// TIA Portal V21 export
// export: Created 2026-10-14T03:08:58.0952126Z, ExportSetting WithDefaults, DisplayName Totally Integrated Automation Portal, DisplayVersion V21, DisplayName STEP 7 Professional, DisplayVersion V21, DisplayName STEP 7 Safety, DisplayVersion V21, DisplayName Tech WebApplication, DisplayVersion V21, DisplayName WinCC Basic/Comfort/Advanced, DisplayVersion V21, DisplayName WinCC Unified, DisplayVersion V21
FUNCTION_BLOCK "FB_5_CIP_Simulation_Graph"   // FB7, GRAPH
VERSION : 0.1
// stored: AcknowledgeErrorsRequired true, AutoNumber true, GraphVersion 6.0, InitialValuesAcquisition false, IsIECCheckEnabled false, LanguageInNetworks LAD, LockOperatingMode false, PermanentILProcessingInMANMode false, SetENOAutomatically false, SkipSteps false, UDAEnableTagReadback false, WithAlarmHandling true
   // inherited from GRAPH_BASE
   VAR
      OFF_SQ_BASE : Bool;
   END_VAR
   VAR_INPUT
      OFF_SQ { ExternalAccessible := 'False'; ExternalVisible := 'False'; ExternalWritable := 'False'} : Bool := false;   // Turn sequence off
      INIT_SQ { ExternalAccessible := 'False'; ExternalVisible := 'False'; ExternalWritable := 'False'} : Bool := false;   // Set sequence to initial state
      ACK_EF { ExternalAccessible := 'False'; ExternalVisible := 'False'; ExternalWritable := 'False'} : Bool := false;   // Acknowledge all errors and faults
      S_PREV { ExternalAccessible := 'False'; ExternalVisible := 'False'; ExternalWritable := 'False'} : Bool := false;   // Output previous step in parameter S_NO
      S_NEXT { ExternalAccessible := 'False'; ExternalVisible := 'False'; ExternalWritable := 'False'} : Bool := false;   // Indicate next step in parameter S_NO
      SW_AUTO { ExternalAccessible := 'False'; ExternalVisible := 'False'; ExternalWritable := 'False'} : Bool := false;   // Automatic mode
      SW_TAP { ExternalAccessible := 'False'; ExternalVisible := 'False'; ExternalWritable := 'False'} : Bool := false;   // Semiautomatic/switch with transition
      SW_TOP { ExternalAccessible := 'False'; ExternalVisible := 'False'; ExternalWritable := 'False'} : Bool := false;   // Semiautomatic/ignore transition
      SW_MAN { ExternalAccessible := 'False'; ExternalVisible := 'False'; ExternalWritable := 'False'} : Bool := false;   // Manual mode
      S_SEL { ExternalAccessible := 'False'; ExternalVisible := 'False'; ExternalWritable := 'False'} : Int := 0;   // Select step to be output to S_NO
      S_ON { ExternalAccessible := 'False'; ExternalVisible := 'False'; ExternalWritable := 'False'} : Bool := false;   // Activate step indicated in S_NO
      S_OFF { ExternalAccessible := 'False'; ExternalVisible := 'False'; ExternalWritable := 'False'} : Bool := false;   // Disable step indicated in S_NO
      T_PUSH { ExternalAccessible := 'False'; ExternalVisible := 'False'; ExternalWritable := 'False'} : Bool := false;   // Enable transition to switch in semi automatic mode
   END_VAR
   VAR_OUTPUT
      S_NO { ExternalAccessible := 'False'; ExternalVisible := 'False'; ExternalWritable := 'False'} : Int := 0;   // Step number
      S_MORE { ExternalAccessible := 'False'; ExternalVisible := 'False'; ExternalWritable := 'False'} : Bool := false;   // More steps are available and can be shown in S_NO
      S_ACTIVE { ExternalAccessible := 'False'; ExternalVisible := 'False'; ExternalWritable := 'False'} : Bool := false;   // Step indicated in S_NO is active
      ERR_FLT { ExternalAccessible := 'False'; ExternalVisible := 'False'; ExternalWritable := 'False'} : Bool := false;   // Interlock or supervision group error
      AUTO_ON { ExternalAccessible := 'False'; ExternalVisible := 'False'; ExternalWritable := 'False'} : Bool := false;   // Automatic mode is active
      TAP_ON { ExternalAccessible := 'False'; ExternalVisible := 'False'; ExternalWritable := 'False'} : Bool := false;   // Semiautomatic mode/step with transition enabled
      TOP_ON { ExternalAccessible := 'False'; ExternalVisible := 'False'; ExternalWritable := 'False'} : Bool := false;   // Semiautomatic mode/ignore transition enabled
      MAN_ON { ExternalAccessible := 'False'; ExternalVisible := 'False'; ExternalWritable := 'False'} : Bool := false;   // Manual mode is active
   END_VAR
   VAR_IN_OUT
      cip : "typeCIP";
      stepInitial : Bool;   // Initial step is active
      step1Active : Bool;   // Step 1 is active
      step2Active : Bool;   // Step 2 is active
      step3Active : Bool;   // Step 3 is active
      step4Active : Bool;   // Step 4 is active
   END_VAR
   VAR
      statTemperature : Real;
      statConcentration : Real;
      statAbnomaly : Real;
   END_VAR
   VAR_TEMP
      tempRet : Int;
      tempRandomFlowrate : Int;
      tempRandomAbnomaly : Real;
   END_VAR
BEGIN
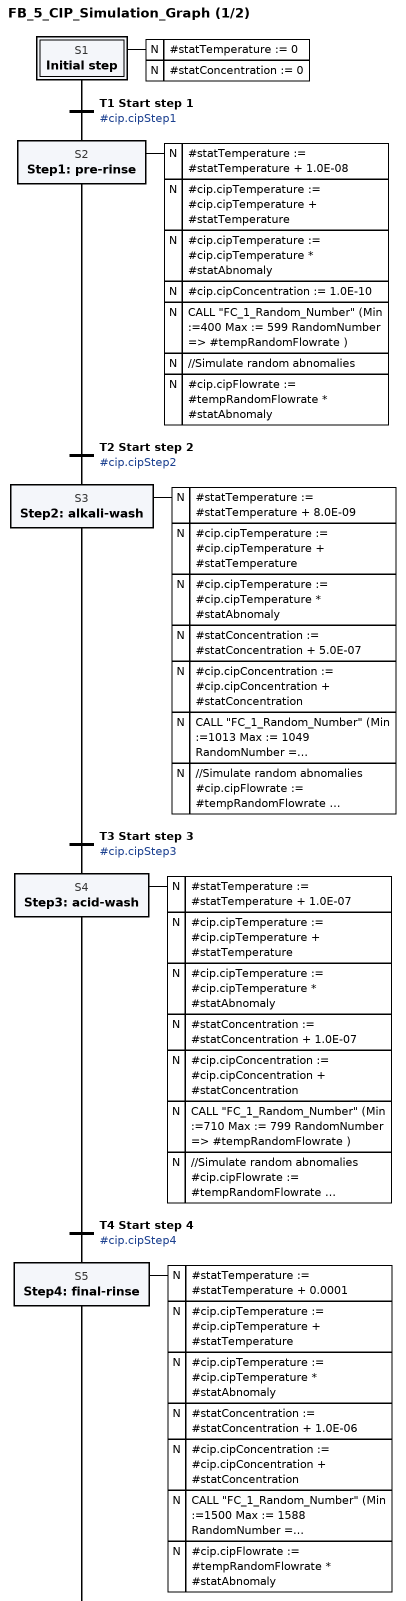
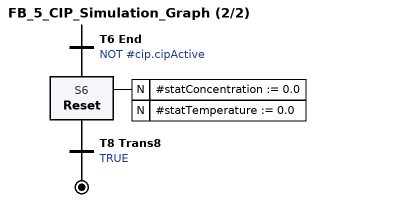
   // permanent pre-instructions
   NETWORK 1
   TITLE = Simulate random abnomalies
      "FC_1_Random_Number"(Min := 70, Max := 100, RandomNumber => #tempRandomAbnomaly);
      #statAbnomaly := #tempRandomAbnomaly / 100.0;

   // sequencer 1
   INITIAL_STEP "Initial step":   // S1, max time T#10S, warning time T#7S
              N    #statTemperature := 0
              N    #statConcentration := 0
   END_STEP
   TRANSITION "Start step 1" FROM "Initial step" TO "Step1: pre-rinse"   // T1
      := #cip.cipStep1;
   END_TRANSITION
   STEP "Step1: pre-rinse":   // S2, max time T#10S, warning time T#7S
              N    #statTemperature := #statTemperature + 1.0E-08
              N    #cip.cipTemperature := #cip.cipTemperature + #statTemperature
              N    #cip.cipTemperature := #cip.cipTemperature * #statAbnomaly
              N    #cip.cipConcentration := 1.0E-10
              N    CALL "FC_1_Random_Number"
                   (Min :=400
                   Max := 599
                   RandomNumber => #tempRandomFlowrate
                   )
                   //Simulate random abnomalies
              N    #cip.cipFlowrate := #tempRandomFlowrate * #statAbnomaly
   END_STEP
   TRANSITION "Start step 2" FROM "Step1: pre-rinse" TO "Step2: alkali-wash"   // T2
      := #cip.cipStep2;
   END_TRANSITION
   STEP "Step2: alkali-wash":   // S3, max time T#10S, warning time T#7S
              N    #statTemperature := #statTemperature + 8.0E-09
              N    #cip.cipTemperature := #cip.cipTemperature + #statTemperature
              N    #cip.cipTemperature := #cip.cipTemperature * #statAbnomaly
              N    #statConcentration := #statConcentration + 5.0E-07
              N    #cip.cipConcentration := #cip.cipConcentration + #statConcentration
              N    CALL "FC_1_Random_Number"
                   (Min :=1013
                   Max := 1049
                   RandomNumber => #tempRandomFlowrate
                   )
              N    //Simulate random abnomalies
                   #cip.cipFlowrate := #tempRandomFlowrate * #statAbnomaly
   END_STEP
   TRANSITION "Start step 3" FROM "Step2: alkali-wash" TO "Step3: acid-wash"   // T3
      := #cip.cipStep3;
   END_TRANSITION
   STEP "Step3: acid-wash":   // S4, max time T#10S, warning time T#7S
              N    #statTemperature := #statTemperature + 1.0E-07
              N    #cip.cipTemperature := #cip.cipTemperature + #statTemperature
              N    #cip.cipTemperature := #cip.cipTemperature * #statAbnomaly
              N    #statConcentration := #statConcentration + 1.0E-07
              N    #cip.cipConcentration := #cip.cipConcentration + #statConcentration
              N    CALL "FC_1_Random_Number"
                   (Min :=710
                   Max := 799
                   RandomNumber => #tempRandomFlowrate
                   )
              N    //Simulate random abnomalies
                   #cip.cipFlowrate := #tempRandomFlowrate * #statAbnomaly
   END_STEP
   TRANSITION "Start step 4" FROM "Step3: acid-wash" TO "Step4: final-rinse"   // T4
      := #cip.cipStep4;
   END_TRANSITION
   STEP "Step4: final-rinse":   // S5, max time T#10S, warning time T#7S
              N    #statTemperature := #statTemperature + 0.0001
              N    #cip.cipTemperature := #cip.cipTemperature + #statTemperature
              N    #cip.cipTemperature := #cip.cipTemperature * #statAbnomaly
              N    #statConcentration := #statConcentration + 1.0E-06
              N    #cip.cipConcentration := #cip.cipConcentration + #statConcentration
              N    CALL "FC_1_Random_Number"
                   (Min :=1500
                   Max := 1588
                   RandomNumber => #tempRandomFlowrate
                   )
              N    #cip.cipFlowrate := #tempRandomFlowrate * #statAbnomaly
   END_STEP
   TRANSITION End FROM "Step4: final-rinse" TO Reset   // T6
      := NOT #cip.cipActive;
   END_TRANSITION
   STEP Reset:   // S6, max time T#10S, warning time T#7S
              N    #statConcentration := 0.0
              N    #statTemperature := 0.0
   END_STEP
   TRANSITION Trans8 FROM Reset TO END   // T8
      := TRUE;
   END_TRANSITION

   // permanent post-instructions
   NETWORK 1
   TITLE = transfer states to output
      #step1Active := #"Step1: pre-rinse".X;
      #step2Active := #"Step2: alkali-wash".X;
      #step3Active := #"Step3: acid-wash".X;
      #step4Active := #"Step4: final-rinse".X;
      #stepInitial := #"Initial step".X;
END_FUNCTION_BLOCK
